INTERFACE I_RoomTempControl

PROPERTY bAlarm : BOOL
GET
END_GET
SET
END_SET
END_PROPERTY

PROPERTY nRoomTemp : REAL
GET
END_GET
END_PROPERTY

END_INTERFACE

(* stored: Version 1.1.0.1
   Itf I_RoomTempControl: Id {7f258d7a-27bc-4e5b-bac9-670543498c63}
   Property bAlarm: Id {098c6b71-9e74-4ee0-94a0-f086b2c06488}
   Get Get: Id {67b7039f-e818-481c-8266-991246e9ffc5}
   Set Set: Id {d33ad352-8510-479d-9e97-c8f1fc4aa2af}
   Property nRoomTemp: Id {e1b4056e-a903-4bcb-85d8-1d188783f658}
   Get Get: Id {c67c22e4-25fc-4bcb-b688-d90eb51c9d53} *)
